(* IEC 61131-3 sources: test/Class/SdiasSDCIMaster (part 3) *)

          TempDataLen := 39;

          InitializeSdoWriteData(Usage:=_SendFunctionCode, ParaIndex:=0, ParaSubIndex:=0, PortSelection:=SIOL_MASTER_PORT_NO, LengthOfData:=TempDataLen, pData:=#TempData[0]);

          sSdoData.eResponseState := t_ReponseState::_SendData;

      //***************************************************************************************************
        t_ReponseState::_SendData,
        t_ReponseState::_Wait4SendResponse,
        t_ReponseState::_GotSendResponse,
        t_ReponseState::_ReadData,
        t_ReponseState::_Wait4ReceiveData,
        t_ReponseState::_GotReceiveData:
          if HandleSdoDataTransfer() = ERROR then
            sSdoData.eAsySSW := _AsyError;
            return;
          end_if;

      //***************************************************************************************************
        t_ReponseState::_GotAllReceiveData:// we enter this step, when we received the answer with the data

          GetSdoReadData(pLength:=#TempDataLen, pData:=#TempData[0]);
          if TempDataLen = 3 then
            // check response data
            if (TempData[0] = (E_FNCID_SETPORTCNFPAR)$USINT) & // check function ID
               (TempData[1] = sSdoData.ActPortSelection)       // check port number
               then

              if (TempData[2] = 0) then // check status code seperately
                // reset response state machine
                sSdoData.eResponseState := t_ReponseState::_PrepareSendData;

                sSdoData.eAsySSW := t_AsySSW::_SwitchToDisableMode;
              else
                // error at return code
                sSdoData.eAsySSW := _AsyError;
                sSdoData.AsyErrorCode := t_SDCIRetCode::SDCI_MicroCtrl_UnexpectedRspData;
                LogError("@503 (SdiasSDCIMaster::AsySSW) Error at status code in answer from µC (_DisablePorts)");
                return;
              end_if;
            else
              // unexpected answer data
              sSdoData.eAsySSW := _AsyError;
              sSdoData.AsyErrorCode := t_SDCIRetCode::SDCI_MicroCtrl_UnexpectedRspData;
              LogError("@0504 (SdiasSDCIMaster::AsySSW) Unexpected data in answer from µC: wrong function ID or port number (_DisablePorts)");
              return;
            end_if;
          else
            // invalid length of answer data
            sSdoData.eAsySSW := _AsyError;
            sSdoData.AsyErrorCode := t_SDCIRetCode::SDCI_MicroCtrl_UnexpectedRspLength;
            LogError("@0505 (SdiasSDCIMaster::AsySSW) Invalid data length in answer from µC (_DisablePorts)");
            return;
          end_if;

      //***************************************************************************************************
      end_case;

//**********************************************************************************************************************************************************
  	t_AsySSW::_SwitchToDisableMode:
      case sSdoData.eResponseState of
      //***************************************************************************************************
        t_ReponseState::_PrepareSendData: // start the sending action
          TempFlags := 0;
          if sSdoData.eAsySSW = t_AsySSW::_SwitchToDisableMode then
  //          TempFlags.Start2Operate := TRUE; // only makes sense if the port is active in SDCI mode
            TempFlags.OperatingMode := TRUE;
          end_if;

          // prepare the sdo buffer
          TempData[0]       := E_FNCID_CNTSTA; // function ID

          // reset the area for all devices before setting for the specific
          _memset(dest:=#TempData[1], usByte:=0, cntr:=SIOL_MAX_PORTS_SUPPORTED * sizeof(TempFlags));

          // activate the disabled mode for the selected port
          TempData[1 + sSdoData.ActPortSelection*sizeof(UINT)]$UINT := TempFlags;

          if TotalMappingWriteSize then
            _memcpy(ptr1:=#TempData[9], ptr2:=#LocalWritePDOBuf[0], cntr:=TotalMappingWriteSize);
          end_if;

          TempDataLen := 9 + TotalMappingWriteSize;

          InitializeSdoWriteData(Usage:=_SendFunctionCode, ParaIndex:=0, ParaSubIndex:=0, PortSelection:=SIOL_MASTER_PORT_NO, LengthOfData:=TempDataLen, pData:=#TempData[0]);

          sSdoData.eResponseState := t_ReponseState::_SendData;

      //***************************************************************************************************
        t_ReponseState::_SendData,
        t_ReponseState::_Wait4SendResponse,
        t_ReponseState::_GotSendResponse,
        t_ReponseState::_ReadData,
        t_ReponseState::_Wait4ReceiveData,
        t_ReponseState::_GotReceiveData:
          if HandleSdoDataTransfer() = ERROR then
            sSdoData.eAsySSW := _AsyError;
            return;
          end_if;

      //***************************************************************************************************
        t_ReponseState::_GotAllReceiveData:// we enter this step, when we received the answer with the data

          GetSdoReadData(pLength:=#TempDataLen, pData:=#TempData[0]);
          if TempDataLen = 9 then
            // check response data
            if (TempData[0] = (E_FNCID_CNTSTA)$USINT) then // check function ID
              // reset response state machine
              sSdoData.eResponseState := t_ReponseState::_PrepareSendData;

              Wait4DeviceDisableStartTime := ops.tAbsolute;

              sSdoData.eAsySSW   := t_AsySSW::_Wait4DisableMode;
            else
              // unexpected answer data
              sSdoData.eAsySSW := _AsyError;
              sSdoData.AsyErrorCode := t_SDCIRetCode::SDCI_MicroCtrl_UnexpectedRspData;
              LogError("@0506 (SdiasSDCIMaster::AsySSW) Unexpected data in answer from µC: wrong function ID or port number (_SwitchToDisableMode)");
              return;
            end_if;
          else
            // invalid length of answer data
            sSdoData.eAsySSW := _AsyError;
            sSdoData.AsyErrorCode := t_SDCIRetCode::SDCI_MicroCtrl_UnexpectedRspLength;
            LogError("@0507 (SdiasSDCIMaster::AsySSW) Invalid data length in answer from µC (_SwitchToDisableMode)");
            return;
          end_if;

      //***************************************************************************************************
      end_case;

//**********************************************************************************************************************************************************
    t_AsySSW::_Wait4DisableMode:
      // if it's a SDCI Portmode, we have to wait for the operating bit to be cleared (maximum time, if it does not get cleared)
      if (aPortInfo[sSdoData.ActPortSelection].CfgPortMode <> _SDCI) |
         ((CyclicInfoTotal.FlagsRdy2OpAndOperating SHR (4+sSdoData.ActPortSelection) AND 1) = FALSE) |
         ((ops.tAbsolute - Wait4DeviceDisableStartTime) > aPortInfo[sSdoData.ActPortSelection].udModeChangeTime) then

        // finished, continue with next step
        if sSdoData.TargetMode = _Inactive then
          // we're on our target state => show it on the class
          sSdoData.eAsySSW   := t_AsySSW::_UpdateClassState;
        else
          // continue setting the new mode
          sSdoData.eAsySSW   := t_AsySSW::_ConfigurePort;
        end_if;
      end_if;

//**********************************************************************************************************************************************************
  	t_AsySSW::_ConfigurePort:
      // if it's a SDCI port, we must wait the time (according to the specification), because some sensors might need it
      if (aPortInfo[sSdoData.ActPortSelection].CfgPortMode = _SDCI) & ((ops.tAbsolute - Wait4DeviceDisableStartTime) < aPortInfo[sSdoData.ActPortSelection].udModeChangeTime) then
        return;
      end_if;

      case sSdoData.eResponseState of
      //***************************************************************************************************
        t_ReponseState::_PrepareSendData: // start the sending action

          // prepare the sdo buffer
          TempData[0]       := E_FNCID_SETPORTCNFPAR; // function ID
          TempData[1]       := sSdoData.ActPortSelection; // port number
          case sSdoData.TargetMode of
          //***************************************************************************************************
            _Inactive:
              TempData[2]       := t_OpModeStates::E_OPMODE_INACTIVE; // operating mode

          //***************************************************************************************************
            _DigitalInput:
              TempData[2]       := t_OpModeStates::E_OPMODE_DI; // operating mode

          //***************************************************************************************************
            _DigitalOutput:
              TempData[2]       := t_OpModeStates::E_OPMODE_DO; // operating mode

          //***************************************************************************************************
            _SDCI:
              TempData[2]       := t_OpModeStates::E_OPMODE_FIXEDMODE; // operating mode

          //***************************************************************************************************
          end_case;

          TempData[3]       := t_PortCycle::E_PORTCYCLE_FIXVAL; // port cycle

          // check if a user override is active
          if aPortInfo[sSdoData.ActPortSelection].OverrideMinCycleTime_us then
            // recalculate cycle time from [µs] to [100µs]
            TempCycleTime     := to_uint(aPortInfo[sSdoData.ActPortSelection].OverrideMinCycleTime_us / 100);
          else
            // recalculate cycle time from [µs] to [100µs]
            TempCycleTime     := to_uint(aPortInfo[sSdoData.ActPortSelection].MinCycleTime_us / 100);
          end_if;

          // make endian swap
          TempCycleTime     := ((TempCycleTime SHR 8) AND 16#FF) OR ((TempCycleTime SHL 8) AND 16#FF00);

          TempData[4]$UINT  := TempCycleTime; // cycle time
          TempData[6]       :=  aPortInfo[sSdoData.ActPortSelection].PdoMapping.ReadDataLength$USINT; // PDConfig LenIn
          TempData[7]       := (aPortInfo[sSdoData.ActPortSelection].PdoMapping.ReadDataStartAddress - SIOL_OFFSET_RT_READ_DATA)$USINT; // PdConfig PosIn
          TempData[8]       := 0; // PdConfig SrcOffsetIn
          TempData[9]       :=  aPortInfo[sSdoData.ActPortSelection].PdoMapping.WriteDataLength$USINT; // PDConfig LenOut
          TempData[10]      := (aPortInfo[sSdoData.ActPortSelection].PdoMapping.WriteDataStartAddress - SIOL_OFFSET_RT_WRITE_DATA)$USINT; // PdConfig PosOut
          TempData[11]      := 0; // PdConfig SrcOffsetOut
          TempData[12]      := (aPortInfo[sSdoData.ActPortSelection].VendorID SHR 8)$USINT; // VendorID
          TempData[13]      :=  aPortInfo[sSdoData.ActPortSelection].VendorID$USINT; // VendorID
          TempData[14]      := (aPortInfo[sSdoData.ActPortSelection].DeviceID SHR 24)$USINT; // DeviceID
          TempData[15]      := (aPortInfo[sSdoData.ActPortSelection].DeviceID SHR 16)$USINT; // DeviceID
          TempData[16]      := (aPortInfo[sSdoData.ActPortSelection].DeviceID SHR  8)$USINT; // DeviceID
          TempData[17]      := (aPortInfo[sSdoData.ActPortSelection].DeviceID       )$USINT; // DeviceID
//          _strcpy(dest:=#TempData[18], src:="0000000000000000"); // serial number as string
          _memset(dest:=#TempData[18], usByte:=0, cntr:=16); // serial number as string
          TempData[34]      := 1; // Inspection level (1 = device and vendor id have to match)
          TempData[35]      := 0; // DS activation state
          TempData[36]      := 0; // DS download enable
          TempData[37]      := 0; // DS upload enable
          TempData[38]      := aPortInfo[sSdoData.ActPortSelection].RevisionID; // revision ID

          TempDataLen := 39;

          InitializeSdoWriteData(Usage:=_SendFunctionCode, ParaIndex:=0, ParaSubIndex:=0, PortSelection:=SIOL_MASTER_PORT_NO, LengthOfData:=TempDataLen, pData:=#TempData[0]);

          sSdoData.eResponseState := t_ReponseState::_SendData;

      //***************************************************************************************************
        t_ReponseState::_SendData,
        t_ReponseState::_Wait4SendResponse,
        t_ReponseState::_GotSendResponse,
        t_ReponseState::_ReadData,
        t_ReponseState::_Wait4ReceiveData,
        t_ReponseState::_GotReceiveData:
          if HandleSdoDataTransfer() = ERROR then
            sSdoData.eAsySSW := _AsyError;
            return;
          end_if;

      //***************************************************************************************************
        t_ReponseState::_GotAllReceiveData:// we enter this step, when we received the answer with the data

          GetSdoReadData(pLength:=#TempDataLen, pData:=#TempData[0]);
          if TempDataLen = 3 then
            // check response data
            if (TempData[0] = (E_FNCID_SETPORTCNFPAR)$USINT) & // check function ID
               (TempData[1] = sSdoData.ActPortSelection)              // check port number
               then

              if (TempData[2] = 0) then // check status code seperately
                // reset response state machine
                sSdoData.eResponseState := t_ReponseState::_PrepareSendData;

                sSdoData.eAsySSW := t_AsySSW::_SwitchToNewMode;
              else
                // error at return code
                sSdoData.eAsySSW := _AsyError;
                sSdoData.AsyErrorCode := t_SDCIRetCode::SDCI_MicroCtrl_UnexpectedRspData;
                LogError("@0508 (SdiasSDCIMaster::AsySSW) Error at status code in answer from µC (_ConfigurePorts)");
                return;
              end_if;
            else
              // unexpected answer data
              sSdoData.eAsySSW := _AsyError;
              sSdoData.AsyErrorCode := t_SDCIRetCode::SDCI_MicroCtrl_UnexpectedRspData;
              LogError("@0509 (SdiasSDCIMaster::AsySSW) Unexpected data in answer from µC: wrong function ID or port number (_ConfigurePorts)");
              return;
            end_if;
          else
            // invalid length of answer data
            sSdoData.eAsySSW := _AsyError;
            sSdoData.AsyErrorCode := t_SDCIRetCode::SDCI_MicroCtrl_UnexpectedRspLength;
            LogError("@050B (SdiasSDCIMaster::AsySSW) Invalid data length in answer from µC  (_ConfigurePorts)");
            return;
          end_if;

      //***************************************************************************************************
      end_case;

//**********************************************************************************************************************************************************
  	t_AsySSW::_SwitchToNewMode:
      case sSdoData.eResponseState of
      //***************************************************************************************************
        t_ReponseState::_PrepareSendData: // start the sending action
          TempFlags := 0;
          TempFlags.Start2Operate := TRUE;
          TempFlags.OperatingMode := TRUE;

          // prepare the sdo buffer
          TempData[0]       := E_FNCID_CNTSTA; // function ID

          // reset the area for all devices before setting for the specific
          _memset(dest:=#TempData[1], usByte:=0, cntr:=SIOL_MAX_PORTS_SUPPORTED * sizeof(TempFlags));

          // activate the new mode for the selected port
          TempData[1 + sSdoData.ActPortSelection*sizeof(UINT)]$UINT := TempFlags;

          if TotalMappingWriteSize then
            _memcpy(ptr1:=#TempData[9], ptr2:=#LocalWritePDOBuf[0], cntr:=TotalMappingWriteSize);
          end_if;

          TempDataLen := 9 + TotalMappingWriteSize;

          InitializeSdoWriteData(Usage:=_SendFunctionCode, ParaIndex:=0, ParaSubIndex:=0, PortSelection:=SIOL_MASTER_PORT_NO, LengthOfData:=TempDataLen, pData:=#TempData[0]);

          sSdoData.eResponseState := t_ReponseState::_SendData;

      //***************************************************************************************************
        t_ReponseState::_SendData,
        t_ReponseState::_Wait4SendResponse,
        t_ReponseState::_GotSendResponse,
        t_ReponseState::_ReadData,
        t_ReponseState::_Wait4ReceiveData,
        t_ReponseState::_GotReceiveData:
          if HandleSdoDataTransfer() = ERROR then
            sSdoData.eAsySSW := _AsyError;
            return;
          end_if;

      //***************************************************************************************************
        t_ReponseState::_GotAllReceiveData:// we enter this step, when we received the answer with the data

          GetSdoReadData(pLength:=#TempDataLen, pData:=#TempData[0]);
          if TempDataLen = 9 then
            // check response data
            if (TempData[0] = (E_FNCID_CNTSTA)$USINT) then // check function ID
              // reset response state machine
              sSdoData.eResponseState := t_ReponseState::_PrepareSendData;

              // remember when we started to wait
              sSdoData.TimeoutStart   := ops.tAbsolute;

              sSdoData.eAsySSW   := t_AsySSW::_Wait4NewMode; // wait until fault or operating
            else
              // unexpected answer data
              sSdoData.eAsySSW := _AsyError;
              sSdoData.AsyErrorCode := t_SDCIRetCode::SDCI_MicroCtrl_UnexpectedRspData;
              LogError("@050C (SdiasSDCIMaster::AsySSW) Unexpected data in answer from µC: wrong function ID or port number (_SwitchToNewMode)");
              return;
            end_if;
          else
            // invalid length of answer data
            sSdoData.eAsySSW := _AsyError;
            sSdoData.AsyErrorCode := t_SDCIRetCode::SDCI_MicroCtrl_UnexpectedRspLength;
            LogError("@050D (SdiasSDCIMaster::AsySSW) Invalid data length in answer from µC (_SwitchToNewMode)");
            return;
          end_if;

      //***************************************************************************************************
      end_case;

//**********************************************************************************************************************************************************
    t_AsySSW::_Wait4NewMode:
      // if mode is not SDCI or operating or fault
      if (sSdoData.TargetMode <> _SDCI) |
         ((CyclicInfoTotal.FlagsRdy2OpAndOperating SHR (4+sSdoData.ActPortSelection) AND 1) = TRUE) |
         ((CyclicInfoTotal.FaultFlags$UINT SHR (sSdoData.ActPortSelection * 4)) AND 16#F) then
        if (sSdoData.TargetMode = _SDCI) & aPortInfo[sSdoData.ActPortSelection].PdoMapping.WriteDataLength then
          // we need to enable the output data also
          sSdoData.eAsySSW   := t_AsySSW::_SetOperateAndPdOutValid;
        else
          // show the class state
          sSdoData.eAsySSW   := t_AsySSW::_UpdateClassState;
        end_if;
      elsif (ops.tAbsolute - sSdoData.TimeoutStart) > SIOL_SDO_RESPONSE_TIMEOUT  then
        sSdoData.eAsySSW := _AsyError;
        sSdoData.AsyErrorCode := t_SDCIRetCode::SDCI_TimeoutInComToMicroCtrl;
        LogError("@0513 (SdiasSDCIMaster::AsySSW) Timeout when waiting for operate when switching the port mode (_Wait4NewMode)");
      end_if;

//**********************************************************************************************************************************************************
  	t_AsySSW::_SetOperateAndPdOutValid:
      case sSdoData.eResponseState of
      //***************************************************************************************************
        t_ReponseState::_PrepareSendData: // start the sending action
          TempFlags := 0;
          TempFlags.Start2Operate := TRUE;
          TempFlags.OperatingMode := TRUE;

          // prepare the sdo buffer
          TempData[0]       := E_FNCID_CNTSTA; // function ID

          TempFlags.PdOutValid := aPortInfo[sSdoData.ActPortSelection].PdoMapping.WriteDataLength <> 0;

          // reset the area for all devices before setting for the specific
          _memset(dest:=#TempData[1], usByte:=0, cntr:=SIOL_MAX_PORTS_SUPPORTED * sizeof(TempFlags));

          TempData[1 + sSdoData.ActPortSelection*sizeof(UINT)]$UINT := TempFlags;

          if TotalMappingWriteSize then
            _memset(dest:=#TempData[9], usByte:=0, cntr:=TotalMappingWriteSize);
          end_if;

          TempDataLen := 9 + TotalMappingWriteSize;

          InitializeSdoWriteData(Usage:=_SendFunctionCode, ParaIndex:=0, ParaSubIndex:=0, PortSelection:=SIOL_MASTER_PORT_NO, LengthOfData:=TempDataLen, pData:=#TempData[0]);

          sSdoData.eResponseState := t_ReponseState::_SendData;

      //***************************************************************************************************
        t_ReponseState::_SendData,
        t_ReponseState::_Wait4SendResponse,
        t_ReponseState::_GotSendResponse,
        t_ReponseState::_ReadData,
        t_ReponseState::_Wait4ReceiveData,
        t_ReponseState::_GotReceiveData:
          if HandleSdoDataTransfer() = ERROR then
            sSdoData.eAsySSW := _AsyError;
            return;
          end_if;

      //***************************************************************************************************
        t_ReponseState::_GotAllReceiveData:// we enter this step, when we received the answer with the data

          GetSdoReadData(pLength:=#TempDataLen, pData:=#TempData[0]);
          if TempDataLen = 9 then
            // check response data
            if (TempData[0] = (E_FNCID_CNTSTA)$USINT) then // check function ID
              // reset response state machine
              sSdoData.eResponseState := t_ReponseState::_PrepareSendData;

              // if the operating flag is cleared we can continue
              TempStateFlags := TempData[1 + sSdoData.ActPortSelection*sizeof(t_StatusFlags)]$t_StatusFlags;

              sSdoData.eAsySSW   := t_AsySSW::_Wait4Operate; // wait until fault or operating
            else
              // unexpected answer data
              sSdoData.eAsySSW := _AsyError;
              sSdoData.AsyErrorCode := t_SDCIRetCode::SDCI_MicroCtrl_UnexpectedRspData;
              LogError("@0515 (SdiasSDCIMaster::AsySSW) Unexpected data in answer from µC: wrong function ID or port number (_ActivatePdOut)");
              return;
            end_if;
          else
            // invalid length of answer data
            sSdoData.eAsySSW := _AsyError;
            sSdoData.AsyErrorCode := t_SDCIRetCode::SDCI_MicroCtrl_UnexpectedRspLength;
            LogError("@0516 (SdiasSDCIMaster::AsySSW) Invalid data length in answer from µC (_ActivatePdOut)");
            return;
          end_if;

      //***************************************************************************************************
      end_case;

  //**********************************************************************************************************************************************************
    t_AsySSW::_Wait4Operate:
      // if operating or fault
      if ((CyclicInfoTotal.FlagsRdy2OpAndOperating SHR (4+sSdoData.ActPortSelection) AND 1) = TRUE) |
         ((CyclicInfoTotal.FaultFlags$UINT SHR (sSdoData.ActPortSelection * 4)) AND 16#F) then

        // show class state
        sSdoData.eAsySSW   := t_AsySSW::_UpdateClassState;
      end_if;

  //**********************************************************************************************************************************************************
    t_AsySSW::_UpdateClassState:
      // if it's a reconnect and the device is not available, we're only here because we wanted to deactivate the port
      if (sSdoData.AsyCmdType = Reconnect) & (aPortInfo[sSdoData.ActPortSelection].PhysicallyAvailable = FALSE) then
        // the object already shows the correct state
      else
        // in all other cases, show the device state at the object

        // save target mode to current mode
        aPortInfo[sSdoData.ActPortSelection].ActPortMode := sSdoData.TargetMode;

        // if there is an object to update
        if aPortInfo[sSdoData.ActPortSelection].pThis then

          // set the command
          MyPara.uiCmd    := CMD_SIOL_DEVICE_INFO_UPDATE;

          // if it's SDCI
          if (aPortInfo[sSdoData.ActPortSelection].ActPortMode = _SDCI) then

            // if there is an IODD file
            if aPortInfo[sSdoData.ActPortSelection].pCfgTable then

              // class state
              if (aPortInfo[sSdoData.ActPortSelection].MinCycleTime_us | aPortInfo[sSdoData.ActPortSelection].OverrideMinCycleTime_us) & aPortInfo[sSdoData.ActPortSelection].VendorID & aPortInfo[sSdoData.ActPortSelection].DeviceID then

                // device available => check if it's the right one
                if (aPortInfo[sSdoData.ActPortSelection].VendorID = aPortInfo[sSdoData.ActPortSelection].pCfgTable^.VendorID) & (aPortInfo[sSdoData.ActPortSelection].DeviceID = aPortInfo[sSdoData.ActPortSelection].pCfgTable^.DeviceID) then
                  // we're good here
                  MyPara.aPara[0] := _ClassOk$DINT;
                  aPortInfo[sSdoData.ActPortSelection].PhysicallyAvailable := TRUE;
                else
                  // wrong device
                  MyPara.aPara[0] := _WrongHardware$DINT;

                  // with this it doesn't get enabled when the fixed mode is set on all ports (doesn't make sense if it's the wrong module)
                  aPortInfo[sSdoData.ActPortSelection].PhysicallyAvailable := FALSE;
                end_if;
              else
                // device not available
                MyPara.aPara[0] := _NoHardware$DINT;

                aPortInfo[sSdoData.ActPortSelection].PhysicallyAvailable := FALSE;
              end_if;
            else
              // no IODD file => any device is ok if one of the Device Infos is available
              if aPortInfo[sSdoData.ActPortSelection].MinCycleTime_us | aPortInfo[sSdoData.ActPortSelection].OverrideMinCycleTime_us | aPortInfo[sSdoData.ActPortSelection].VendorID | aPortInfo[sSdoData.ActPortSelection].DeviceID then
                // we're good here
                MyPara.aPara[0] := _ClassOk$DINT;
                aPortInfo[sSdoData.ActPortSelection].PhysicallyAvailable := TRUE;
              else
                // no device infos available
                MyPara.aPara[0] := _NoHardware$DINT;

                aPortInfo[sSdoData.ActPortSelection].PhysicallyAvailable := FALSE;
              end_if;
            end_if;

            // vendor ID
            MyPara.aPara[1] := aPortInfo[sSdoData.ActPortSelection].VendorID;

            // device ID
            MyPara.aPara[2] := aPortInfo[sSdoData.ActPortSelection].DeviceID$DINT;

            // minimum cycle time
            // check if a user override is active
            if aPortInfo[sSdoData.ActPortSelection].OverrideMinCycleTime_us then
              MyPara.aPara[3] := aPortInfo[sSdoData.ActPortSelection].OverrideMinCycleTime_us$DINT;
            else
              MyPara.aPara[3] := aPortInfo[sSdoData.ActPortSelection].MinCycleTime_us$DINT;
            end_if;

            // actual port mode
            MyPara.aPara[4] := t_SDCIPortMode::_SDCI;

            if aPortInfo[sSdoData.ActPortSelection].Required & (MyPara.aPara[0] <> _NotInitialized$DINT) then
              // show required error on SDCI device
              MyPara.aPara[0] := _RequiredError$DINT;
              aPortInfo[sSdoData.ActPortSelection].pThis^.NewInst(#MyPara, #MyResult);

              SetRequiredError();
            else
              aPortInfo[sSdoData.ActPortSelection].pThis^.NewInst(#MyPara, #MyResult);
            end_if;

          else
            // it's always ok here
            MyPara.aPara[0] := _ClassOk$DINT;
            aPortInfo[sSdoData.ActPortSelection].PhysicallyAvailable := TRUE;

            // vendor ID
            MyPara.aPara[1] := aPortInfo[sSdoData.ActPortSelection].VendorID;

            // device ID
            MyPara.aPara[2] := aPortInfo[sSdoData.ActPortSelection].DeviceID$DINT;

            // minimum cycle time
            // check if a user override is active
            if aPortInfo[sSdoData.ActPortSelection].OverrideMinCycleTime_us then
              MyPara.aPara[3] := aPortInfo[sSdoData.ActPortSelection].OverrideMinCycleTime_us$DINT;
            else
              MyPara.aPara[3] := aPortInfo[sSdoData.ActPortSelection].MinCycleTime_us$DINT;
            end_if;

            // actual port mode is already valid here (no further changes on the setting of this port)
            MyPara.aPara[4] := aPortInfo[sSdoData.ActPortSelection].ActPortMode$DINT;

            aPortInfo[sSdoData.ActPortSelection].pThis^.NewInst(#MyPara, #MyResult);
          end_if;
        end_if;
      end_if;

      if sSdoData.AsyCmdType = DelayedEnable then
        // remove the bit from the current port from the ToDo-list and go to the next port
        DelayedEnablePorts := DelayedEnablePorts SHR 1;
        sSdoData.ActPortSelection += 1;

        // check if there are more modules to enable
        sSdoData.eAsySSW  := t_AsySSW::_StartDelayedEnable;
      else
        //last reconnect of one port
        sAutoConnectVars.udLastReconnectTry := ops.tAbsolute;
        // we're finished
        sSdoData.eAsySSW := t_AsySSW::_Finished;
      end_if;

  //**********************************************************************************************************************************************************
  t_AsySSW::_Finished:
      sSdoData.eAsySSW  := t_AsySSW::_Idle;
      sSdoData.AsyState := t_SDCIRetCode::SDCI_Ready_Ok;

      // Handle Asy Callback
      if sSdoData.pCallBackThis & sSdoData.pCallBackFun then
        HandleSDOCallback();
      end_if;

      // Unlock SDO Channel
      sigclib_atomic_setU32(pValue:=#sSdoData.DataLock, value:= SSDCIM_SDO_UNLOCK);

  //**********************************************************************************************************************************************************
    t_AsySSW::_AsyError:
      sSdoData.eAsySSW  := t_AsySSW::_Idle;

      // use the stored error code
      sSdoData.AsyState := sSdoData.AsyErrorCode;

      // Handle Asy Callback
      if sSdoData.pCallBackThis & sSdoData.pCallBackFun then
        HandleSDOCallback();
      end_if;

      // Unlock SDO Channel
      sigclib_atomic_setU32(pValue:=#sSdoData.DataLock, value:= SSDCIM_SDO_UNLOCK);

  //**********************************************************************************************************************************************************
  end_case;

#ifdef SIOL_ENABLE_DEBUG_LOGGING
  if sSdoData.eAsySSW <> OldAsyStep then
    AsyStepTimes[OldAsyStep$DINT] := ops.tAbsolute;
    OldAsyStep := sSdoData.eAsySSW;
  end_if;
#pragma message("RamAnd 31.01.2017 10:41 \ testweise die Zeit der einzelnen Steps messen")
#endif

END_FUNCTION

FUNCTION SdiasSDCIMaster::ChangeModeIsPossible
	VAR_INPUT
		TargetPort 	: USINT;
		TargetMode 	: SdiasSDCIMaster::t_SDCIPortMode;
	END_VAR
	VAR_OUTPUT
		ChangeIsPossible 	: BOOL;
	END_VAR

  if (TargetMode = _DigitalInput) & (aPortInfo[TargetPort].PdoMapping.ReadDataLength = 0) then
    // cannot change to digital input mode if there is no possibility to transfer the input value
    ChangeIsPossible := FALSE;
  elsif (TargetMode = _DigitalOutput) & (aPortInfo[TargetPort].PdoMapping.WriteDataLength = 0) then
    // cannot change to digital output mode if there is no possibility to transfer the output value
    ChangeIsPossible := FALSE;
  else
    ChangeIsPossible := TRUE;
  end_if;

END_FUNCTION

FUNCTION SdiasSDCIMaster::InitTheModule
	VAR_OUTPUT
		eModuleInitState 	: iprStates;
	END_VAR
  VAR
  	TempData            : ARRAY [0..SIOL_MAX_SDO_DATA_SIZE-1] OF USINT;
    TempDataLen         : USINT;
    TempFlags           : t_ControlFlags;
    TempStateFlags      : t_StatusFlags;
    i                   : DINT;
  	MyPara              : CmdStruct;
    MyResult            : results;
    TempCycleTime       : UINT;
    SDCIPortAvailable   : BOOL;
    DigStartUpAvailable : BOOL;
  END_VAR

  // if the returncode isn't changed to ERROR or READY, we return busy
  eModuleInitState := BUSY;

  case sSdoData.eInitSSW of
//**********************************************************************************************************************************************************
  	t_InitSSW::_InitVariables:

      // reset asy state machine variables
      sSdoData.AsyState         := t_SDCIRetCode::SDCI_Ready_Ok;
      sSdoData.eAsySSW          := _Idle;

      // prepare initialisation
      sSdoData.ActPortSelection := 0;
      sSdoData.eResponseState   := t_ReponseState::_ReadData;
      sSdoData.eInitSSW         := t_InitSSW::_GetFwInfo;

      //get value for waittime between reconnects
      WaitTimeReconnect := WaitTimeReconnect.Read();
      if WaitTimeReconnect > SIOL_MINIMUM_WAIT4RECONNECT_TIME*2 then
        WaitTimeReconnect := SIOL_MINIMUM_WAIT4RECONNECT_TIME*2;
      end_if;

//**********************************************************************************************************************************************************
    t_InitSSW::_GetFwInfo:

      case sSdoData.eResponseState of
        //***************************************************************************************************
          t_ReponseState::_ReadData:// we enter this step to start the read access

            sSdoData.ActDataSize       := sizeof(t_FirmwareInfo);
            sSdoData.pActData          := #FwInfo;

            StartReadSDO(hOffset:=SIOL_OFFSET_INFO_FOR_PLC, usLength:=sSdoData.ActDataSize, eCommand:=SDIAS_SDO_CMD_MEM_READ);
            sSdoData.TimeoutStart   := ops.tAbsolute;
            sSdoData.eResponseState := t_ReponseState::_Wait4ReceiveData;

        //***************************************************************************************************
          t_ReponseState::_Wait4ReceiveData:// we wait for the read data
            if (ops.tAbsolute - sSdoData.TimeoutStart) > SIOL_SDO_TIMEOUT then
              LogError("@0517 (SdiasSDCIMaster::InitTheModule) Timeout at reading firmware info from module");
              sSdoData.eInitSSW := _Error;
              return;
            end_if;

        //***************************************************************************************************
          t_ReponseState::_GotReceiveData:// we enter this step, when we received the answer with the data
            // receivedata in the right place => continue with the next step

            // show the version at the server if the crc is correct
            if (FwInfo.LengthOfData = 0) | (CheckSum_16(pData:=#FwInfo.Data.Version, uiDataLength:=FwInfo.LengthOfData, uiCRCStart:=16#FFFF) <> FwInfo.CRC) then
              if FwInfo.LengthOfData = 0 then
                LogError("@0518 (SdiasSDCIMaster::InitTheModule) No firmware available!");
                sSdoData.eInitSSW := _Error;
                return;
              else
                LogError("@0519 (SdiasSDCIMaster::InitTheModule) Incorrect checksum of info from µC detected!");
              end_if;
            end_if;

            FirmwareVersion := FwInfo.Data.Version;

            sSdoData.eResponseState   := t_ReponseState::_ReadData;
            sSdoData.eInitSSW         := t_InitSSW::_GetActMessageCnt;

        //***************************************************************************************************
      end_case;

//**********************************************************************************************************************************************************
    t_InitSSW::_GetActMessageCnt:

      case sSdoData.eResponseState of

        //***************************************************************************************************
          t_ReponseState::_ReadData:// we enter this step to start the read access

            sSdoData.ActDataSize       := sizeof(t_ServiceDataArea.wo_MessageCnt);
            sSdoData.pActData          := #sSdoData.SdoWriteData.wo_MessageCnt;

            StartReadSDO(hOffset:=SIOL_OFFSET_SERVICE_DATA_AREA + t_ServiceDataArea.wo_MessageCnt, usLength:=sSdoData.ActDataSize, eCommand:=SDIAS_SDO_CMD_MEM_READ);
            sSdoData.TimeoutStart   := ops.tAbsolute;
            sSdoData.eResponseState := t_ReponseState::_Wait4ReceiveData;

        //***************************************************************************************************
          t_ReponseState::_Wait4ReceiveData:// we wait for the read data
            if (ops.tAbsolute - sSdoData.TimeoutStart) > SIOL_SDO_TIMEOUT then
              LogError("@051A (SdiasSDCIMaster::InitTheModule) Timeout at reading actual message counter from module");
              sSdoData.eInitSSW := _Error;
              return;
            end_if;

        //***************************************************************************************************
          t_ReponseState::_GotReceiveData:// we enter this step, when we received the answer with the data
            // receivedata in the right place => continue with the next step

            // take the read counter as first write counter (continue counting after reset/run of the PLC)
            sSdoData.SdoReadData.ro_MessageCnt := sSdoData.SdoWriteData.wo_MessageCnt;

            sSdoData.eResponseState   := t_ReponseState::_PrepareSendData;
            sSdoData.eInitSSW         := t_InitSSW::_Set24VSupplyOn;

        //***************************************************************************************************
      end_case;

//**********************************************************************************************************************************************************
    t_InitSSW::_Set24VSupplyOn:
      case sSdoData.eResponseState of
      //***************************************************************************************************
        t_ReponseState::_PrepareSendData: // start the sending action

          // prepare the sdo buffer
          TempData[0]       := E_FNCID_SWITCHON; // function ID
          TempData[1]       := sSdoData.ActPortSelection; // port number

          TempDataLen := 2;

          InitializeSdoWriteData(Usage:=_SendFunctionCode, ParaIndex:=0, ParaSubIndex:=0, PortSelection:=SIOL_MASTER_PORT_NO, LengthOfData:=TempDataLen, pData:=#TempData[0]);

          sSdoData.eResponseState := t_ReponseState::_SendData;

      //***************************************************************************************************
        t_ReponseState::_SendData,
        t_ReponseState::_Wait4SendResponse,
        t_ReponseState::_GotSendResponse,
        t_ReponseState::_ReadData,
        t_ReponseState::_Wait4ReceiveData,
        t_ReponseState::_GotReceiveData:
          if HandleSdoDataTransfer() = ERROR then
            sSdoData.eInitSSW := _Error;
            return;
          end_if;

      //***************************************************************************************************
        t_ReponseState::_GotAllReceiveData:// we enter this step, when we received the answer with the data

          GetSdoReadData(pLength:=#TempDataLen, pData:=#TempData[0]);
          if TempDataLen = 2 then
            // check response data
            if (TempData[0] = (E_FNCID_SWITCHON)$USINT) then // check function ID
              if (TempData[1] = 0) then                                     // check status code seperately
                // reset response state machine
                sSdoData.eResponseState := t_ReponseState::_PrepareSendData;

                // already the last port?
                if sSdoData.ActPortSelection = (SIOL_MAX_PORTS_SUPPORTED-1) then
                  // finished, continue with next step
                  sSdoData.ActPortSelection := 0;

                  sSdoData.eInitSSW := t_InitSSW::_DisablePorts;
                else
                  // repeat the step with the next port
                  sSdoData.ActPortSelection += 1;
                end_if;
              else
                // error at return code
                LogError("@051B (SdiasSDCIMaster::InitTheModule) Error at status code in answer from µC (_Set24VSupplyOn)");
                sSdoData.eInitSSW := _Error;
                return;
              end_if;
            else
              // unexpected answer data
              LogError("@051C (SdiasSDCIMaster::InitTheModule) Unexpected data in answer from µC: wrong function ID  (_Set24VSupplyOn)");
              sSdoData.eInitSSW := _Error;
              return;
            end_if;
          else
            // invalid length of answer data
            LogError("@051D (SdiasSDCIMaster::InitTheModule) Invalid data length in answer from µC  (_Set24VSupplyOn)");
            sSdoData.eInitSSW := _Error;
            return;
          end_if;

      //***************************************************************************************************
      end_case;

//**********************************************************************************************************************************************************
  	t_InitSSW::_DisablePorts:
      case sSdoData.eResponseState of
      //***************************************************************************************************
        t_ReponseState::_PrepareSendData: // start the sending action

          // prepare the sdo buffer
          TempData[0]       := E_FNCID_SETPORTCNFPAR; // function ID
          TempData[1]       := sSdoData.ActPortSelection; // port number
          TempData[2]       := t_OpModeStates::E_OPMODE_INACTIVE; // operating mode
          TempData[3]       := t_PortCycle::E_PORTCYCLE_FREERN; // port cycle
          TempData[4]$UINT  := 0; // cycle time
          TempData[6]       :=  aPortInfo[sSdoData.ActPortSelection].PdoMapping.ReadDataLength$USINT; // PDConfig LenIn
          TempData[7]       := (aPortInfo[sSdoData.ActPortSelection].PdoMapping.ReadDataStartAddress - SIOL_OFFSET_RT_READ_DATA)$USINT; // PdConfig PosIn
          TempData[8]       := 0; // PdConfig SrcOffsetIn
          TempData[9]       :=  aPortInfo[sSdoData.ActPortSelection].PdoMapping.WriteDataLength$USINT; // PDConfig LenOut
          TempData[10]      := (aPortInfo[sSdoData.ActPortSelection].PdoMapping.WriteDataStartAddress - SIOL_OFFSET_RT_WRITE_DATA)$USINT; // PdConfig PosOut
          TempData[11]      := 0; // PdConfig SrcOffsetOut
          TempData[12]$UINT := 0; // VendorID
          TempData[14]$UDINT:= 0; // DeviceID
//          _strcpy(dest:=#TempData[18], src:="0000000000000000"); // serial number as string
          _memset(dest:=#TempData[18], usByte:=0, cntr:=16); // serial number as string
          TempData[34]      := 0; // Inspection level
          TempData[35]      := 0; // DS activation state
          TempData[36]      := 0; // DS download enable
          TempData[37]      := 0; // DS upload enable
          TempData[38]      := 16#11; // revision ID (v1.1 should work with both device types, v1.0 doesn't work with v1.1 devices)

          TempDataLen := 39;

          InitializeSdoWriteData(Usage:=_SendFunctionCode, ParaIndex:=0, ParaSubIndex:=0, PortSelection:=SIOL_MASTER_PORT_NO, LengthOfData:=TempDataLen, pData:=#TempData[0]);

          sSdoData.eResponseState := t_ReponseState::_SendData;

      //***************************************************************************************************
        t_ReponseState::_SendData,
        t_ReponseState::_Wait4SendResponse,
        t_ReponseState::_GotSendResponse,
        t_ReponseState::_ReadData,
        t_ReponseState::_Wait4ReceiveData,
        t_ReponseState::_GotReceiveData:
          if HandleSdoDataTransfer() = ERROR then
            sSdoData.eInitSSW := _Error;
            return;
          end_if;

      //***************************************************************************************************
        t_ReponseState::_GotAllReceiveData:// we enter this step, when we received the answer with the data

          GetSdoReadData(pLength:=#TempDataLen, pData:=#TempData[0]);
          if TempDataLen = 3 then
            // check response data
            if (TempData[0] = (E_FNCID_SETPORTCNFPAR)$USINT) & // check function ID
               (TempData[1] = sSdoData.ActPortSelection)              // check port number
               then

              if (TempData[2] = 0) then // check status code seperately
                // reset response state machine
                sSdoData.eResponseState := t_ReponseState::_PrepareSendData;

                // already the last port?
                if sSdoData.ActPortSelection = (SIOL_MAX_PORTS_SUPPORTED-1) then
                  // finished, continue with next step
                  sSdoData.ActPortSelection := 0;
                  sSdoData.eInitSSW := t_InitSSW::_SwitchToDisableMode;
                else
                  // repeat the steps with the next port
                  sSdoData.ActPortSelection += 1;
                end_if;
              else
                // error at return code
                LogError("@0503 (SdiasSDCIMaster::InitTheModule) Error at status code in answer from µC (_DisablePorts)");
                sSdoData.eInitSSW := _Error;
                return;
              end_if;
            else
              // unexpected answer data
              LogError("@0504 (SdiasSDCIMaster::InitTheModule) Unexpected data in answer from µC: wrong function ID or port number (_DisablePorts)");
              sSdoData.eInitSSW := _Error;
              return;
            end_if;
          else
            // invalid length of answer data
            LogError("@0505 (SdiasSDCIMaster::InitTheModule) Invalid data length in answer from µC (_DisablePorts)");
            sSdoData.eInitSSW := _Error;
            return;
          end_if;

      //***************************************************************************************************
      end_case;

//**********************************************************************************************************************************************************
  	t_InitSSW::_SwitchToDisableMode,
    t_InitSSW::_Wait4DisableMode:
      case sSdoData.eResponseState of
      //***************************************************************************************************
        t_ReponseState::_PrepareSendData: // start the sending action
          TempFlags := 0;
          if sSdoData.eInitSSW = t_InitSSW::_SwitchToDisableMode then
  //          TempFlags.Start2Operate := TRUE; // only makes sense if the port is active in SDCI mode
            TempFlags.OperatingMode := TRUE;
          end_if;

          // prepare the sdo buffer
          TempData[0]       := E_FNCID_CNTSTA; // function ID
          for i:= 0 to SIOL_MAX_PORTS_SUPPORTED-1 do
            // activate the disabled mode for all ports
            TempData[1 + i*sizeof(UINT)]$UINT := TempFlags;
          end_for;

          if TotalMappingWriteSize then
            _memset(dest:=#TempData[9], usByte:=0, cntr:=TotalMappingWriteSize);
          end_if;

          TempDataLen := 9 + TotalMappingWriteSize;

          InitializeSdoWriteData(Usage:=_SendFunctionCode, ParaIndex:=0, ParaSubIndex:=0, PortSelection:=SIOL_MASTER_PORT_NO, LengthOfData:=TempDataLen, pData:=#TempData[0]);

          sSdoData.eResponseState := t_ReponseState::_SendData;

      //***************************************************************************************************
        t_ReponseState::_SendData,
        t_ReponseState::_Wait4SendResponse,
        t_ReponseState::_GotSendResponse,
        t_ReponseState::_ReadData,
        t_ReponseState::_Wait4ReceiveData,
        t_ReponseState::_GotReceiveData:
          if HandleSdoDataTransfer() = ERROR then
            sSdoData.eInitSSW := _Error;
            return;
          end_if;

      //***************************************************************************************************
        t_ReponseState::_GotAllReceiveData:// we enter this step, when we received the answer with the data

          GetSdoReadData(pLength:=#TempDataLen, pData:=#TempData[0]);
          if TempDataLen = 9 then
            // check response data
            if (TempData[0] = (E_FNCID_CNTSTA)$USINT) then // check function ID
              // reset response state machine
              sSdoData.eResponseState := t_ReponseState::_PrepareSendData;

              // if the operating flags are cleared we can continue
              for i:= 0 to SIOL_MAX_PORTS_SUPPORTED-1 do
                TempStateFlags := TempData[1 + i*sizeof(t_StatusFlags)]$t_StatusFlags;

                // if any operating bit is still set => go to wait for disabled
                if TempStateFlags.Operating = TRUE then

                  // set the time mark the first time we send the command to not wait unnecessary
                  if sSdoData.eInitSSW = t_InitSSW::_SwitchToDisableMode then
                    Wait4DeviceDisableStartTime := ops.tAbsolute;
                  end_if;

                  sSdoData.eInitSSW   := t_InitSSW::_Wait4DisableMode;

                  return;
                end_if;
              end_for;

              // finished, continue with next step
              sSdoData.eInitSSW   := t_InitSSW::_ConfigurePorts;
            else
              // unexpected answer data
              LogError("@0506 (SdiasSDCIMaster::InitTheModule) Unexpected data in answer from µC: wrong function ID or port number (_SwitchToDisableMode)");
              sSdoData.eInitSSW := _Error;
              return;
            end_if;
          else
            // invalid length of answer data
            LogError("@0507 (SdiasSDCIMaster::InitTheModule) Invalid data length in answer from µC (_SwitchToDisableMode)");
            sSdoData.eInitSSW := _Error;
            return;
          end_if;

      //***************************************************************************************************
      end_case;

//**********************************************************************************************************************************************************
  	t_InitSSW::_ConfigurePorts:
      // if it's a SDCI port, we must wait the time (according to the specification), because some sensors might need it
      if (aPortInfo[sSdoData.ActPortSelection].CfgPortMode = _SDCI) & ((ops.tAbsolute - Wait4DeviceDisableStartTime) < aPortInfo[sSdoData.ActPortSelection].udModeChangeTime) then
        return;
      end_if;

      case sSdoData.eResponseState of
      //***************************************************************************************************
        t_ReponseState::_PrepareSendData: // start the sending action

          // prepare the sdo buffer
          TempData[0]       := E_FNCID_SETPORTCNFPAR; // function ID
          TempData[1]       := sSdoData.ActPortSelection; // port number
          case aPortInfo[sSdoData.ActPortSelection].CfgPortMode of
          //***************************************************************************************************
            _Inactive:
              TempData[2]       := t_OpModeStates::E_OPMODE_INACTIVE; // operating mode

          //***************************************************************************************************
            _DigitalInput:
              TempData[2]       := t_OpModeStates::E_OPMODE_DI; // operating mode

          //***************************************************************************************************
            _DigitalOutput:
              TempData[2]       := t_OpModeStates::E_OPMODE_DO; // operating mode

          //***************************************************************************************************
            _SDCI:
              TempData[2]       := t_OpModeStates::E_OPMODE_SCANMODE; // operating mode

          //***************************************************************************************************
          end_case;

          TempData[3]       := t_PortCycle::E_PORTCYCLE_FREERN; // port cycle
          TempData[4]$UINT  := 0; // cycle time
          TempData[6]       :=  aPortInfo[sSdoData.ActPortSelection].PdoMapping.ReadDataLength$USINT; // PDConfig LenIn
          TempData[7]       := (aPortInfo[sSdoData.ActPortSelection].PdoMapping.ReadDataStartAddress - SIOL_OFFSET_RT_READ_DATA)$USINT; // PdConfig PosIn
          TempData[8]       := 0; // PdConfig SrcOffsetIn
          TempData[9]       :=  aPortInfo[sSdoData.ActPortSelection].PdoMapping.WriteDataLength$USINT; // PDConfig LenOut
          TempData[10]      := (aPortInfo[sSdoData.ActPortSelection].PdoMapping.WriteDataStartAddress - SIOL_OFFSET_RT_WRITE_DATA)$USINT; // PdConfig PosOut
          TempData[11]      := 0; // PdConfig SrcOffsetOut
          TempData[12]$UINT := 0; // VendorID
          TempData[14]$UDINT:= 0; // DeviceID
//          _strcpy(dest:=#TempData[18], src:="0000000000000000"); // serial number as string
          _memset(dest:=#TempData[18], usByte:=0, cntr:=16); // serial number as string
          TempData[34]      := 0; // Inspection level (0 = don't care about vendor or device id)
          TempData[35]      := 0; // DS activation state
          TempData[36]      := 0; // DS download enable
          TempData[37]      := 0; // DS upload enable
          TempData[38]      := 16#11; // revision ID (v1.1 should work with both device types, v1.0 doesn't work with v1.1 devices)

          TempDataLen := 39;

          InitializeSdoWriteData(Usage:=_SendFunctionCode, ParaIndex:=0, ParaSubIndex:=0, PortSelection:=SIOL_MASTER_PORT_NO, LengthOfData:=TempDataLen, pData:=#TempData[0]);

          sSdoData.eResponseState := t_ReponseState::_SendData;

      //***************************************************************************************************
        t_ReponseState::_SendData,
        t_ReponseState::_Wait4SendResponse,
        t_ReponseState::_GotSendResponse,
        t_ReponseState::_ReadData,
        t_ReponseState::_Wait4ReceiveData,
        t_ReponseState::_GotReceiveData:
          if HandleSdoDataTransfer() = ERROR then
            sSdoData.eInitSSW := _Error;
            return;
          end_if;

      //***************************************************************************************************
        t_ReponseState::_GotAllReceiveData:// we enter this step, when we received the answer with the data

          GetSdoReadData(pLength:=#TempDataLen, pData:=#TempData[0]);
          if TempDataLen = 3 then
            // check response data
            if (TempData[0] = (E_FNCID_SETPORTCNFPAR)$USINT) & // check function ID
               (TempData[1] = sSdoData.ActPortSelection)              // check port number
               then

              if (TempData[2] = 0) then // check status code seperately
                // reset response state machine
                sSdoData.eResponseState := t_ReponseState::_PrepareSendData;

                // already the last port?
                if sSdoData.ActPortSelection = (SIOL_MAX_PORTS_SUPPORTED-1) then
                  // finished, continue with next step
                  sSdoData.ActPortSelection := 0;
                  sSdoData.eInitSSW := t_InitSSW::_EnableMasterServices;
                else
                  // repeat the steps with the next port
                  sSdoData.ActPortSelection += 1;
                end_if;
              else
                // error at return code
                LogError("@0508 (SdiasSDCIMaster::InitTheModule) Error at status code in answer from µC (_ConfigurePorts)");
                sSdoData.eInitSSW := _Error;
                return;
              end_if;
            else
              // unexpected answer data
              LogError("@0509 (SdiasSDCIMaster::InitTheModule) Unexpected data in answer from µC: wrong function ID or port number (_ConfigurePorts)");
              sSdoData.eInitSSW := _Error;
              return;
            end_if;
          else
            // invalid length of answer data
            LogError("@050B (SdiasSDCIMaster::InitTheModule) Invalid data length in answer from µC  (_ConfigurePorts)");
            sSdoData.eInitSSW := _Error;
            return;
          end_if;

      //***************************************************************************************************
      end_case;

//**********************************************************************************************************************************************************
  	t_InitSSW::_EnableMasterServices:
      case sSdoData.eResponseState of
      //***************************************************************************************************
        t_ReponseState::_PrepareSendData: // start the sending action
          TempFlags := 0;
          TempFlags.OdStart       := TRUE;
          TempFlags.DuStart       := TRUE;
          TempFlags.PdStart       := TRUE;

          // prepare the sdo buffer
          TempData[0]       := E_FNCID_CNTSTA; // function ID
          for i:= 0 to SIOL_MAX_PORTS_SUPPORTED-1 do
            // activate the master services for all ports
            TempData[1 + i*sizeof(UINT)]$UINT := TempFlags;
          end_for;

          if TotalMappingWriteSize then
            _memset(dest:=#TempData[9], usByte:=0, cntr:=TotalMappingWriteSize);
          end_if;

          TempDataLen := 9 + TotalMappingWriteSize;

          InitializeSdoWriteData(Usage:=_SendFunctionCode, ParaIndex:=0, ParaSubIndex:=0, PortSelection:=SIOL_MASTER_PORT_NO, LengthOfData:=TempDataLen, pData:=#TempData[0]);

          sSdoData.eResponseState := t_ReponseState::_SendData;

      //***************************************************************************************************
        t_ReponseState::_SendData,
        t_ReponseState::_Wait4SendResponse,
        t_ReponseState::_GotSendResponse,
        t_ReponseState::_ReadData,
        t_ReponseState::_Wait4ReceiveData,
        t_ReponseState::_GotReceiveData:
          if HandleSdoDataTransfer() = ERROR then
            sSdoData.eInitSSW := _Error;
            return;
          end_if;

      //***************************************************************************************************
        t_ReponseState::_GotAllReceiveData:// we enter this step, when we received the answer with the data

          GetSdoReadData(pLength:=#TempDataLen, pData:=#TempData[0]);
          if TempDataLen = 9 then
            // check response data
            if (TempData[0] = (E_FNCID_CNTSTA)$USINT) then // check function ID
              // reset response state machine
              sSdoData.eResponseState := t_ReponseState::_PrepareSendData;

              for i:= 0 to SIOL_MAX_PORTS_SUPPORTED-1 do
                if aPortInfo[i].pThis then
                  aPortInfo[i].PhysicallyAvailable := TRUE;
                else
                  aPortInfo[i].PhysicallyAvailable := FALSE;
                end_if;
              end_for;

              // continue with next step
              sSdoData.eInitSSW := t_InitSSW::_SwitchToNewMode;
            else
              // unexpected answer data
              LogError("@051F (SdiasSDCIMaster::InitTheModule) Unexpected data in answer from µC: wrong function ID or port number (_EnableMasterServices)");
              sSdoData.eInitSSW := _Error;
              return;
            end_if;
          else
            // invalid length of answer data
            LogError("@0520 (SdiasSDCIMaster::InitTheModule) Invalid data length in answer from µC (_EnableMasterServices)");
            sSdoData.eInitSSW := _Error;
            return;
          end_if;

      //***************************************************************************************************
      end_case;

//**********************************************************************************************************************************************************

  	t_InitSSW::_SwitchToNewMode,
    t_InitSSW::_Wait4NewMode:
      case sSdoData.eResponseState of
      //***************************************************************************************************
        t_ReponseState::_PrepareSendData: // start the sending action
          TempFlags := 0;
          if sSdoData.eInitSSW = t_InitSSW::_SwitchToNewMode then
            TempFlags.Start2Operate := TRUE;
            TempFlags.OperatingMode := TRUE;
          end_if;

          // prepare the sdo buffer
          TempData[0]       := E_FNCID_CNTSTA; // function ID
          for i:= 0 to SIOL_MAX_PORTS_SUPPORTED-1 do

            // activate the disabled mode for all ports
            TempData[1 + i*sizeof(UINT)]$UINT := TempFlags;

          end_for;

          if TotalMappingWriteSize then
            _memset(dest:=#TempData[9], usByte:=0, cntr:=TotalMappingWriteSize);
          end_if;

          TempDataLen := 9 + TotalMappingWriteSize;

          InitializeSdoWriteData(Usage:=_SendFunctionCode, ParaIndex:=0, ParaSubIndex:=0, PortSelection:=SIOL_MASTER_PORT_NO, LengthOfData:=TempDataLen, pData:=#TempData[0]);

          sSdoData.eResponseState := t_ReponseState::_SendData;

      //***************************************************************************************************
        t_ReponseState::_SendData,
        t_ReponseState::_Wait4SendResponse,
        t_ReponseState::_GotSendResponse,
        t_ReponseState::_ReadData,
        t_ReponseState::_Wait4ReceiveData,
        t_ReponseState::_GotReceiveData:
          if HandleSdoDataTransfer() = ERROR then
            sSdoData.eInitSSW := _Error;
            return;
          end_if;

      //***************************************************************************************************
        t_ReponseState::_GotAllReceiveData:// we enter this step, when we received the answer with the data

          GetSdoReadData(pLength:=#TempDataLen, pData:=#TempData[0]);
          if TempDataLen = 9 then

            // reset response state machine
            sSdoData.eResponseState := t_ReponseState::_PrepareSendData;

            // check response data
            if (TempData[0] = (E_FNCID_CNTSTA)$USINT) then // check function ID

              // if the operating flags are cleared we can continue
              for i:= 0 to SIOL_MAX_PORTS_SUPPORTED-1 do
                TempStateFlags := TempData[1 + i*sizeof(t_StatusFlags)]$t_StatusFlags;

                // if any operating bit is not set and there is also no fault => go to wait again
                if (aPortInfo[i].CfgPortMode = _SDCI) & (TempStateFlags.Operating = FALSE) &
                   ((TempStateFlags AND 16#F000) = 0) then // no fault
                  sSdoData.eInitSSW   := t_InitSSW::_Wait4NewMode; // wait until fault or operating
                  return;
                end_if;
              end_for;

              // finished, continue with next step
              sSdoData.eInitSSW   := t_InitSSW::_GetDeviceInfos;
            else
              // unexpected answer data
              LogError("@050C (SdiasSDCIMaster::InitTheModule) Unexpected data in answer from µC: wrong function ID or port number (_SwitchToNewMode)");
              sSdoData.eInitSSW := _Error;
              return;
            end_if;
          else
            // invalid length of answer data
            LogError("@050D (SdiasSDCIMaster::InitTheModule) Invalid data length in answer from µC (_SwitchToNewMode)");
            sSdoData.eInitSSW := _Error;
            return;
          end_if;

      //***************************************************************************************************
      end_case;

//**********************************************************************************************************************************************************
    t_InitSSW::_GetDeviceInfos:

      case sSdoData.eResponseState of
      //***************************************************************************************************
        t_ReponseState::_PrepareSendData: // start the sending action
          if aPortInfo[sSdoData.ActPortSelection].CfgPortMode = _SDCI then

            // read direct parameter page 1 (device info)
            InitializeSdoWriteData(Usage:=_ReadParaData, ParaIndex:=0, ParaSubIndex:=0, PortSelection:=sSdoData.ActPortSelection, LengthOfData:=0, pData:=NIL);

            sSdoData.eResponseState := t_ReponseState::_SendData;

          else
            // already the last port?
            if sSdoData.ActPortSelection = (SIOL_MAX_PORTS_SUPPORTED-1) then
              // finished, continue with next step
              sSdoData.ActPortSelection := 0;

              sSdoData.eInitSSW := t_InitSSW::_UpdateDeviceObjInfo;
            else
              // repeat the step with the next port
              sSdoData.ActPortSelection += 1;
            end_if;
          end_if;

      //***************************************************************************************************
        t_ReponseState::_SendData,
        t_ReponseState::_Wait4SendResponse,
        t_ReponseState::_GotSendResponse,
        t_ReponseState::_ReadData,
        t_ReponseState::_Wait4ReceiveData,
        t_ReponseState::_GotReceiveData:
          if HandleSdoDataTransfer() = ERROR then
            sSdoData.eInitSSW := _Error;
            return;
          end_if;

      //***************************************************************************************************
        t_ReponseState::_GotAllReceiveData:// we enter this step, when we received the answer with the data

          // reset response state machine
          sSdoData.eResponseState := t_ReponseState::_PrepareSendData;

          GetSdoReadData(pLength:=#TempDataLen, pData:=#TempData[0]);
          if (sSdoData.SdoReadData.ro_RetCode = _ServiceNotAvailable) | (TempDataLen = 0) then
            // maybe the port is not connected => select next port (after this if block)
            aPortInfo[sSdoData.ActPortSelection].PhysicallyAvailable := FALSE;

          else
#ifdef SIOL_ENABLE_DEBUG_LOGGING
if TempData$t_DeviceInfoAnswer.ProcessDataIn <> aPortInfo[sSdoData.ActPortSelection].PdoMapping.ReadDataBitLength then
  LogValue("@DBG (SdiasSDCIMaster::InitTheModule) Info: Configured bit size of read PDO 0x{0} does not match the expected size from the module 0x{1}. SDCI Port 0x{2}", udValue:=aPortInfo[sSdoData.ActPortSelection].PdoMapping.ReadDataBitLength, udValue2:=TempData$t_DeviceInfoAnswer.ProcessDataIn, udValue3:=sSdoData.ActPortSelection);
end_if;
if TempData$t_DeviceInfoAnswer.ProcessDataOut <> aPortInfo[sSdoData.ActPortSelection].PdoMapping.WriteDataBitLength then
  LogValue("@DBG (SdiasSDCIMaster::InitTheModule) Info: Configured bit size of write PDO 0x{0} does not match the expected size from the module 0x{1}. SDCI Port 0x{2}", udValue:=aPortInfo[sSdoData.ActPortSelection].PdoMapping.WriteDataBitLength, udValue2:=TempData$t_DeviceInfoAnswer.ProcessDataOut, udValue3:=sSdoData.ActPortSelection);
end_if;
#endif

            // MIN CYCLE TIME
            case TempData$t_DeviceInfoAnswer.MinCycleTime SHR 6 of
              0: // base of  100µs (Multiplier x time base)
                aPortInfo[sSdoData.ActPortSelection].MinCycleTime_us :=  100 * (TempData$t_DeviceInfoAnswer.MinCycleTime AND 16#3F);

              1: // base of  400µs (Multiplier x time base) +  6400µs
                aPortInfo[sSdoData.ActPortSelection].MinCycleTime_us :=  400 * (TempData$t_DeviceInfoAnswer.MinCycleTime AND 16#3F) +  6400;

              2: // base of 1600µs (Multiplier x time base) + 32000µs
                aPortInfo[sSdoData.ActPortSelection].MinCycleTime_us := 1600 * (TempData$t_DeviceInfoAnswer.MinCycleTime AND 16#3F) + 32000;

              3: // this is reserved for future use
                LogError("@050E (SdiasSDCIMaster::InitTheModule) Invalid time base 3 received at minimum cycle time of device (_GetDeviceInfos)");
                sSdoData.eInitSSW := _Error;
                return;
            end_case;

            // VENDOR ID
            aPortInfo[sSdoData.ActPortSelection].VendorID := TempData$t_DeviceInfoAnswer.VendorIdLsb OR (TempData$t_DeviceInfoAnswer.VendorIdMsb SHL 8);

            // DEVICE ID
            aPortInfo[sSdoData.ActPortSelection].DeviceID := TempData$t_DeviceInfoAnswer.DeviceIdLsb OR (TempData$t_DeviceInfoAnswer.DeviceIdMiddleByte SHL 8) OR (TempData$t_DeviceInfoAnswer.DeviceIdMsb SHL 16);

            // Revision ID
            aPortInfo[sSdoData.ActPortSelection].RevisionID := TempData$t_DeviceInfoAnswer.RevisionID;

            aPortInfo[sSdoData.ActPortSelection].aDeviceInfo$t_DeviceInfoAnswer := TempData$t_DeviceInfoAnswer;
          end_if;

          // already the last port?
          if sSdoData.ActPortSelection = (SIOL_MAX_PORTS_SUPPORTED-1) then
            // finished, continue with next step
            sSdoData.ActPortSelection := 0;

            sSdoData.eInitSSW := t_InitSSW::_UpdateDeviceObjInfo;
          else
            // repeat the step with the next port
            sSdoData.ActPortSelection += 1;
          end_if;

      //***************************************************************************************************
      end_case;

//**********************************************************************************************************************************************************
    t_InitSSW::_UpdateDeviceObjInfo:

      // if the SDIAS bus is too fast for the SDCI master
      if (udBusTime/1000) < SIOL_MINIMUM_MASTER_CYCLE_TIME then
        // go to the lowest possible value that is a multiple of the bus time
        if SIOL_MINIMUM_MASTER_CYCLE_TIME MOD (udBusTime/1000) then
          // if there is a rest => add 1 to the multiplier
          CycleTime := (udBusTime / 1000)$UINT * ((SIOL_MINIMUM_MASTER_CYCLE_TIME / (udBusTime / 1000)$UINT) + 1);
        else
          // otherwise use the bustime directly to get to the minimum master cycle time
//          CycleTime := (udBusTime / 1000)$UINT * ((SIOL_MINIMUM_MASTER_CYCLE_TIME / (udBusTime / 1000)$UINT)    );
          CycleTime := SIOL_MINIMUM_MASTER_CYCLE_TIME;
        end_if;
      else
        // otherwise take the SDIAS bus time
        CycleTime := (udBusTime / 1000)$UINT;
      end_if;

      SDCIPortAvailable := FALSE;

      // the same command for all objects
      MyPara.uiCmd    := CMD_SIOL_DEVICE_INFO_UPDATE;

      // show the info at the objects and also set the class state server
      for i := 0 to SIOL_MAX_PORTS_SUPPORTED-1 do
        // reset act parameter number for next init step
        aPortInfo[i].ActParaNo := 0;

        // if there is an object to update
        if aPortInfo[i].pThis then

          // if it's SDCI
          if (aPortInfo[i].CfgPortMode = _SDCI) then

            SDCIPortAvailable := TRUE;

            // if there is an IODD file
            if aPortInfo[i].pCfgTable then
              // class state
              if (aPortInfo[i].MinCycleTime_us | aPortInfo[i].OverrideMinCycleTime_us) & aPortInfo[i].VendorID & aPortInfo[i].DeviceID then

                // device available => check if it's the right one
                if (aPortInfo[i].VendorID = aPortInfo[i].pCfgTable^.VendorID) & (aPortInfo[i].DeviceID = aPortInfo[i].pCfgTable^.DeviceID) then
                  // show that we are still initializing
                  MyPara.aPara[0] := _NotInitialized$DINT;
                else
                  // wrong device
                  MyPara.aPara[0] := _WrongHardware$DINT;

                  // with this it doesn't get enabled when the fixed mode is set on all ports (doesn't make sense if it's the wrong module)
                  aPortInfo[i].PhysicallyAvailable := FALSE;
                end_if;
              else
                // device not available
                MyPara.aPara[0] := _NoHardware$DINT;

                aPortInfo[i].PhysicallyAvailable := FALSE;
              end_if;
            else
              // no IODD file => any device is ok if one of the Device Infos is available
              if aPortInfo[i].MinCycleTime_us | aPortInfo[i].OverrideMinCycleTime_us | aPortInfo[i].VendorID | aPortInfo[i].DeviceID then
                // show that we are still initializing
                MyPara.aPara[0] := _NotInitialized$DINT;
              else
                // no device infos available
                MyPara.aPara[0] := _NoHardware$DINT;

                aPortInfo[i].PhysicallyAvailable := FALSE;
              end_if;
            end_if;

            // vendor ID
            MyPara.aPara[1] := aPortInfo[i].VendorID;

            // device ID
            MyPara.aPara[2] := aPortInfo[i].DeviceID$DINT;

            // minimum cycle time
            // check if a user override is active
            if aPortInfo[i].OverrideMinCycleTime_us then
              MyPara.aPara[3] := aPortInfo[i].OverrideMinCycleTime_us$DINT;
            else
              MyPara.aPara[3] := aPortInfo[i].MinCycleTime_us$DINT;
            end_if;

            // actual port mode (still Inactive during initialisation)
            MyPara.aPara[4] := t_SDCIPortMode::_Inactive;

            if aPortInfo[i].Required & (MyPara.aPara[0] <> _NotInitialized$DINT) then
              // show required error on SDCI device
              MyPara.aPara[0] := _RequiredError$DINT;
              aPortInfo[i].pThis^.NewInst(#MyPara, #MyResult);

              SetRequiredError();
            else
              aPortInfo[i].pThis^.NewInst(#MyPara, #MyResult);
            end_if;

          elsif (aPortInfo[i].CfgPortMode = _DigitalInput) | (aPortInfo[i].CfgPortMode = _DigitalOutput) then
            // it's always ok here
            MyPara.aPara[0] := _ClassOk$DINT;

            // we're in the desired mode
            aPortInfo[i].ActPortMode := aPortInfo[i].CfgPortMode;

            // the extra info does not exist here
            MyPara.aPara[1] := 0;
            MyPara.aPara[2] := 0;
            MyPara.aPara[3] := 0;

            // actual port mode is already valid here (no further changes on the setting of this port)
            MyPara.aPara[4] := aPortInfo[i].ActPortMode$DINT;

            aPortInfo[i].pThis^.NewInst(#MyPara, #MyResult);
          end_if;
        end_if;
      end_for;

      if SDCIPortAvailable then
          sSdoData.eInitSSW := t_InitSSW::_CheckDownloadParameters;

        DownloadTimeStart := ops.tAbsolute;

        // if the first pointer is not valid, skip until we find a valid pointer
        if aPortInfo[sSdoData.ActPortSelection].pActPara = NIL then
          if SelectNextDownloadPara() = FALSE then
            // no download parameters available

            sSdoData.ActPortSelection := 0;

            // go to next step
            sSdoData.eInitSSW := t_InitSSW::_DisableSdciPorts;
            // reset response state machine
            sSdoData.eResponseState := t_ReponseState::_PrepareSendData;
          end_if;
        end_if;
      else
        DelayedEnablePorts := 0;

        // no SDCI ports available => skip switching off/on and downloading parameters
        sSdoData.eInitSSW := t_InitSSW::_SetCycleTimes;
      end_if;

//**********************************************************************************************************************************************************
    t_InitSSW::_CheckDownloadParameters:

      case sSdoData.eResponseState of
      //***************************************************************************************************
        t_ReponseState::_PrepareSendData: // start the sending action

          // get the details to write the parameter
          if aPortInfo[sSdoData.ActPortSelection].pActPara then

            if aPortInfo[sSdoData.ActPortSelection].pActPara^.AccessType = t_ParaAccessType::wo then
              // Do not read write only parameters and write the parameter directly
              sSdoData.eInitSSW := t_InitSSW::_DownloadParameters;
            else
              // read the parameter first (to check if it already matches the desired value)
              InitializeSdoWriteData(Usage:=_ReadParaData, ParaIndex:=aPortInfo[sSdoData.ActPortSelection].pActPara^.ParaID$UINT, ParaSubIndex:=aPortInfo[sSdoData.ActPortSelection].pActPara^.ParaSubID$USINT, PortSelection:=sSdoData.ActPortSelection, LengthOfData:=0, pData:=NIL);

              sSdoData.eResponseState := t_ReponseState::_SendData;
            end_if;

          end_if;

      //***************************************************************************************************
        t_ReponseState::_SendData,
        t_ReponseState::_Wait4SendResponse,
        t_ReponseState::_GotSendResponse,
        t_ReponseState::_ReadData,
        t_ReponseState::_Wait4ReceiveData,
        t_ReponseState::_GotReceiveData:
          if HandleSdoDataTransfer() = ERROR then
            sSdoData.eInitSSW := _Error;
            return;
          end_if;

      //***************************************************************************************************
        t_ReponseState::_GotAllReceiveData:// we enter this step, when we received the answer with the data

          // extend the post init time by the reaction time of the µC (otherwise we would exceed the timeout of the post init if there are many parameters)
          ExtendPostInitTime(AdditionalTime:=ops.tAbsolute - sSdoData.ResponseTimeoutStart);

          // reset response state machine
          sSdoData.eResponseState := t_ReponseState::_PrepareSendData;

          // check response data
          if (sSdoData.SdoReadData.ro_RetCode = _FwOk) then // check returncode

            // check if the value matches our init value
            GetSdoReadData( pLength       := #TempDataLen
                          , pData         := #TempData[0]
                          , bDoEndianSwap := CheckEndianSwapNeeded( pParaInfo     := aPortInfo[sSdoData.ActPortSelection].pActPara
                                                                  , PortSelection := sSdoData.ActPortSelection) );

            // if it's a string, we add the termination 0 to the uploaded data (for the comparison), because we also have it in the table
            if aPortInfo[sSdoData.ActPortSelection].pActPara^.DataType = _Text then
              TempData[TempDataLen] := 0;
              TempDataLen += 1;
            end_if;

            if (aPortInfo[sSdoData.ActPortSelection].pActPara^.DataLength = TempDataLen) then
              if _memcmp(ptr1:=#TempData[0], ptr2:=aPortInfo[sSdoData.ActPortSelection].pActPara + sizeof(t_ConfigTablePara), cntr:=TempDataLen) = 0 then
                // value match => no download necessary
#ifdef SIOL_ENABLE_DEBUG_LOGGING
LogValue("@DBG (SdiasSDCIMaster::InitTheModule) Value and length match already, no download needed. ParameterIndex: {0}, ParameterSubIndex: {1}", udValue:=aPortInfo[sSdoData.ActPortSelection].pActPara^.ParaID, udValue2:=aPortInfo[sSdoData.ActPortSelection].pActPara^.ParaSubID);
#endif
              else

                // it's not the same value => download the parameter
                sSdoData.eInitSSW := t_InitSSW::_DownloadParameters;

#ifdef SIOL_ENABLE_DEBUG_LOGGING
LogValue("@DBG (SdiasSDCIMaster::InitTheModule) Value mismatch => download new value. ParameterIndex: {0}, ParameterSubIndex: {1}", udValue:=aPortInfo[sSdoData.ActPortSelection].pActPara^.ParaID, udValue2:=aPortInfo[sSdoData.ActPortSelection].pActPara^.ParaSubID);
#endif

                // skip selecting the next parameter, because we need to send the current parameter in the downloadparameters step
                return;
              end_if;
            else
              // length mismatch

              // if it's a string, we send the new value
              if aPortInfo[sSdoData.ActPortSelection].pActPara^.DataType = _Text then

                // it's not the same value => download the parameter
                sSdoData.eInitSSW := t_InitSSW::_DownloadParameters;

#ifdef SIOL_ENABLE_DEBUG_LOGGING
LogValue("@DBG (SdiasSDCIMaster::InitTheModule) Length mismatch at string => download new value. ParameterIndex: {0}, ParameterSubIndex: {1}", udValue:=aPortInfo[sSdoData.ActPortSelection].pActPara^.ParaID, udValue2:=aPortInfo[sSdoData.ActPortSelection].pActPara^.ParaSubID);
#endif

                // skip selecting the next parameter, because we need to send the current parameter in the downloadparameters step
                return;
              else
                LogValue("@050F (SdiasSDCIMaster::InitTheModule) Length mismatch (type is not string) => value not downloaded. ParameterIndex: {0}, ParameterSubIndex: {1}", udValue:=aPortInfo[sSdoData.ActPortSelection].pActPara^.ParaID, udValue2:=aPortInfo[sSdoData.ActPortSelection].pActPara^.ParaSubID);
              end_if;
            end_if;

            if SelectNextDownloadPara() = FALSE then
              // no more download parameters available

              sSdoData.ActPortSelection := 0;

              // go to next step
              sSdoData.eInitSSW := t_InitSSW::_DisableSdciPorts;
            end_if;
          else
            if (sSdoData.SdoReadData.ro_RetCode = _ApplicationError) then
              // if it's an application error, we also have an error code
              LogValue("@0510 (SdiasSDCIMaster::InitTheModule) Error at reading parameter(_CheckDownloadParameters). ParameterIndex: {0}, ParameterSubIndex: {1}, ErrorCode: {2}", udValue:=aPortInfo[sSdoData.ActPortSelection].pActPara^.ParaID, udValue2:=aPortInfo[sSdoData.ActPortSelection].pActPara^.ParaSubID, udValue3:=sSdoData.SdoReadData.aData[230]$HINT);
            else
              LogValue("@0510 (SdiasSDCIMaster::InitTheModule) Error at reading parameter(_CheckDownloadParameters). ParameterIndex: {0}, ParameterSubIndex: {1}", udValue:=aPortInfo[sSdoData.ActPortSelection].pActPara^.ParaID, udValue2:=aPortInfo[sSdoData.ActPortSelection].pActPara^.ParaSubID);
            end_if;

            // continue with the next parameter
            if SelectNextDownloadPara() = FALSE then
              // no more download parameters available

              sSdoData.ActPortSelection := 0;

              // go to next step
              sSdoData.eInitSSW := t_InitSSW::_DisableSdciPorts;
            end_if;
          end_if;

      //***************************************************************************************************
      end_case;

//**********************************************************************************************************************************************************
    t_InitSSW::_DownloadParameters:

      case sSdoData.eResponseState of
      //***************************************************************************************************
        t_ReponseState::_PrepareSendData: // start the sending action

          // get the details to write the parameter
          if aPortInfo[sSdoData.ActPortSelection].pActPara then

            // prepare everything to send the parameter
            TempDataLen := aPortInfo[sSdoData.ActPortSelection].pActPara^.DataLength;
            _memcpy(ptr1:=#TempData[0], ptr2:=aPortInfo[sSdoData.ActPortSelection].pActPara + sizeof(t_ConfigTablePara), cntr:=TempDataLen);

            InitializeSdoWriteData( Usage         := _WriteParaData
                                  , ParaIndex     := aPortInfo[sSdoData.ActPortSelection].pActPara^.ParaID$UINT
                                  , ParaSubIndex  := aPortInfo[sSdoData.ActPortSelection].pActPara^.ParaSubID$USINT
                                  , PortSelection := sSdoData.ActPortSelection
                                  , LengthOfData  := TempDataLen
                                  , pData         := #TempData[0]
                                  , pParaInfo     := aPortInfo[sSdoData.ActPortSelection].pActPara);

            sSdoData.eResponseState := t_ReponseState::_SendData;
          else
            sSdoData.eInitSSW := _Error;
            LogError("@0521 (SdiasSDCIMaster::InitTheModule) Conditions for parameter download not met. No valid parameter pointer!");
            return;
          end_if;

      //***************************************************************************************************
        t_ReponseState::_SendData,
        t_ReponseState::_Wait4SendResponse,
        t_ReponseState::_GotSendResponse,
        t_ReponseState::_ReadData,
        t_ReponseState::_Wait4ReceiveData,
        t_ReponseState::_GotReceiveData:
          if HandleSdoDataTransfer() = ERROR then
            sSdoData.eInitSSW := _Error;
            return;
          end_if;

      //***************************************************************************************************
        t_ReponseState::_GotAllReceiveData:// we enter this step, when we received the answer with the data

          // extend the post init time by the reaction time of the µC (otherwise we would exceed the timeout of the post init if there are many parameters)
          ExtendPostInitTime(AdditionalTime:=ops.tAbsolute - sSdoData.ResponseTimeoutStart);

          // in general we go back to check the next parameter (unless there are no more parameters)
          sSdoData.eInitSSW := t_InitSSW::_CheckDownloadParameters;

          // reset response state machine
          sSdoData.eResponseState := t_ReponseState::_PrepareSendData;

          // check response data
          if (sSdoData.SdoReadData.ro_RetCode = _FwOk) then // check returncode

#ifdef SIOL_ENABLE_DEBUG_LOGGING
LogValue("@DBG (SdiasSDCIMaster::InitTheModule) Successfully downloaded parameter (_DownloadParameters). ParameterIndex: {0}, ParameterSubIndex: {1}", udValue:=aPortInfo[sSdoData.ActPortSelection].pActPara^.ParaID, udValue2:=aPortInfo[sSdoData.ActPortSelection].pActPara^.ParaSubID);
#endif

          elsif (sSdoData.SdoReadData.ro_RetCode = _ApplicationError) then
            // if it's an application error, we also have an error code
            LogValue("@0512 (SdiasSDCIMaster::InitTheModule) Error at writing parameter(_DownloadParameters). ParameterIndex: {0}, ParameterSubIndex: {1}, ErrorCode: {2}", udValue:=aPortInfo[sSdoData.ActPortSelection].pActPara^.ParaID, udValue2:=aPortInfo[sSdoData.ActPortSelection].pActPara^.ParaSubID, udValue3:=sSdoData.SdoReadData.aData[230]$HINT);
          else
            LogValue("@0512 (SdiasSDCIMaster::InitTheModule) Error at writing parameter(_DownloadParameters). ParameterIndex: {0}, ParameterSubIndex: {1}", udValue:=aPortInfo[sSdoData.ActPortSelection].pActPara^.ParaID, udValue2:=aPortInfo[sSdoData.ActPortSelection].pActPara^.ParaSubID);
          end_if;

          // select the next parameter
          if SelectNextDownloadPara() = FALSE then
            // no more download parameters available

            sSdoData.ActPortSelection := 0;

            // go to next step
            sSdoData.eInitSSW := t_InitSSW::_DisableSdciPorts;

          end_if;

      //***************************************************************************************************
      end_case;

//**********************************************************************************************************************************************************
  	t_InitSSW::_DisableSdciPorts:
      case sSdoData.eResponseState of
      //***************************************************************************************************
        t_ReponseState::_PrepareSendData: // start the sending action

          // only if the port is of type SDCI
          if aPortInfo[sSdoData.ActPortSelection].CfgPortMode = _SDCI then
            // prepare the sdo buffer
            TempData[0]       := E_FNCID_SETPORTCNFPAR; // function ID
            TempData[1]       := sSdoData.ActPortSelection; // port number
            TempData[2]       := t_OpModeStates::E_OPMODE_INACTIVE; // operating mode
            TempData[3]       := t_PortCycle::E_PORTCYCLE_FREERN; // port cycle
            TempData[4]$UINT  := 0; // cycle time
            TempData[6]       :=  aPortInfo[sSdoData.ActPortSelection].PdoMapping.ReadDataLength$USINT; // PDConfig LenIn
            TempData[7]       := (aPortInfo[sSdoData.ActPortSelection].PdoMapping.ReadDataStartAddress - SIOL_OFFSET_RT_READ_DATA)$USINT; // PdConfig PosIn
            TempData[8]       := 0; // PdConfig SrcOffsetIn
            TempData[9]       :=  aPortInfo[sSdoData.ActPortSelection].PdoMapping.WriteDataLength$USINT; // PDConfig LenOut
            TempData[10]      := (aPortInfo[sSdoData.ActPortSelection].PdoMapping.WriteDataStartAddress - SIOL_OFFSET_RT_WRITE_DATA)$USINT; // PdConfig PosOut
            TempData[11]      := 0; // PdConfig SrcOffsetOut
            TempData[12]$UINT := 0; // VendorID
            TempData[14]$UDINT:= 0; // DeviceID
  //          _strcpy(dest:=#TempData[18], src:="0000000000000000"); // serial number as string
            _memset(dest:=#TempData[18], usByte:=0, cntr:=16); // serial number as string
            TempData[34]      := 0; // Inspection level
            TempData[35]      := 0; // DS activation state
            TempData[36]      := 0; // DS download enable
            TempData[37]      := 0; // DS upload enable
            TempData[38]      := 16#11; // revision ID (v1.1 should work with both device types, v1.0 doesn't work with v1.1 devices)

            TempDataLen := 39;

            InitializeSdoWriteData(Usage:=_SendFunctionCode, ParaIndex:=0, ParaSubIndex:=0, PortSelection:=SIOL_MASTER_PORT_NO, LengthOfData:=TempDataLen, pData:=#TempData[0]);

            sSdoData.eResponseState := t_ReponseState::_SendData;
          else
            // already the last port?
            if sSdoData.ActPortSelection = (SIOL_MAX_PORTS_SUPPORTED-1) then
              // finished, continue with next step
              sSdoData.ActPortSelection := 0;

              sSdoData.eInitSSW := t_InitSSW::_SwitchToDisableMode2;

            else
              // repeat the step with the next port
              sSdoData.ActPortSelection += 1;
            end_if;
          end_if;

      //***************************************************************************************************
        t_ReponseState::_SendData,
        t_ReponseState::_Wait4SendResponse,
        t_ReponseState::_GotSendResponse,
        t_ReponseState::_ReadData,
        t_ReponseState::_Wait4ReceiveData,
        t_ReponseState::_GotReceiveData:
          if HandleSdoDataTransfer() = ERROR then
            sSdoData.eInitSSW := _Error;
            return;
          end_if;

      //***************************************************************************************************
        t_ReponseState::_GotAllReceiveData:// we enter this step, when we received the answer with the data

          GetSdoReadData(pLength:=#TempDataLen, pData:=#TempData[0]);
          if TempDataLen = 3 then
            // check response data
            if (TempData[0] = (E_FNCID_SETPORTCNFPAR)$USINT) & // check function ID
               (TempData[1] = sSdoData.ActPortSelection)              // check port number
               then

              if (TempData[2] = 0) then // check status code seperately
                // reset response state machine
                sSdoData.eResponseState := t_ReponseState::_PrepareSendData;

                // already the last port?
                if sSdoData.ActPortSelection = (SIOL_MAX_PORTS_SUPPORTED-1) then
                  // finished, continue with next step
                  sSdoData.ActPortSelection := 0;
                  sSdoData.eInitSSW := t_InitSSW::_SwitchToDisableMode2;
                else
                  // repeat the steps with the next port
                  sSdoData.ActPortSelection += 1;
                end_if;
              else
                // error at return code
                LogError("@0522 (SdiasSDCIMaster::InitTheModule) Error at status code in answer from µC (_DisableSdciPorts)");
                sSdoData.eInitSSW := _Error;
                return;
              end_if;
            else
              // unexpected answer data
              LogError("@0523 (SdiasSDCIMaster::InitTheModule) Unexpected data in answer from µC: wrong function ID or port number (_DisableSdciPorts)");
              sSdoData.eInitSSW := _Error;
              return;
            end_if;
          else
            // invalid length of answer data
            LogError("@0524 (SdiasSDCIMaster::InitTheModule) Invalid data length in answer from µC (_DisableSdciPorts)");
            sSdoData.eInitSSW := _Error;
            return;
          end_if;

          // reset response state machine
          sSdoData.eResponseState := t_ReponseState::_PrepareSendData;

      //***************************************************************************************************
      end_case;

//**********************************************************************************************************************************************************
  	t_InitSSW::_SwitchToDisableMode2,
    t_InitSSW::_Wait4DisableMode2:
      case sSdoData.eResponseState of
      //***************************************************************************************************
        t_ReponseState::_PrepareSendData: // start the sending action
          TempFlags := 0;
          if sSdoData.eInitSSW = t_InitSSW::_SwitchToDisableMode2 then
  //          TempFlags.Start2Operate := TRUE; // only makes sense if the port is active in SDCI mode
            TempFlags.OperatingMode := TRUE;

            Wait4DeviceDisableStartTime := ops.tAbsolute;
          end_if;

          // prepare the sdo buffer
          TempData[0]       := E_FNCID_CNTSTA; // function ID
          for i:= 0 to SIOL_MAX_PORTS_SUPPORTED-1 do
            // activate the disabled mode for all SDCI ports
            if aPortInfo[i].CfgPortMode = _SDCI then
              TempData[1 + i*sizeof(UINT)]$UINT := TempFlags;
            else
              TempData[1 + i*sizeof(UINT)]$UINT := 0;
            end_if;
          end_for;

          if TotalMappingWriteSize then
            _memset(dest:=#TempData[9], usByte:=0, cntr:=TotalMappingWriteSize);
          end_if;

          TempDataLen := 9 + TotalMappingWriteSize;

          InitializeSdoWriteData(Usage:=_SendFunctionCode, ParaIndex:=0, ParaSubIndex:=0, PortSelection:=SIOL_MASTER_PORT_NO, LengthOfData:=TempDataLen, pData:=#TempData[0]);

          sSdoData.eResponseState := t_ReponseState::_SendData;

      //***************************************************************************************************
        t_ReponseState::_SendData,
        t_ReponseState::_Wait4SendResponse,
        t_ReponseState::_GotSendResponse,
        t_ReponseState::_ReadData,
        t_ReponseState::_Wait4ReceiveData,
        t_ReponseState::_GotReceiveData:
          if HandleSdoDataTransfer() = ERROR then
            sSdoData.eInitSSW := _Error;
            return;
          end_if;

      //***************************************************************************************************
        t_ReponseState::_GotAllReceiveData:// we enter this step, when we received the answer with the data
